// TIA Portal V20 export
// export: Created 2026-10-19T18:36:12.7338711Z, ExportSetting WithDefaults, DisplayName Totally Integrated Automation Portal, DisplayVersion V20 Update 6, DisplayName TIA Portal Openness, DisplayVersion V20 Update 6, DisplayName TIA Portal Version Control Interface, DisplayVersion V20 Update 6, DisplayName SINAMICS Startdrive Advanced, DisplayVersion V20 SP1, DisplayName SINAMICS Startdrive G130, G150, S120, S150, SINAMICS MV, G220, S200, S210, DisplayVersion V20 SP1, DisplayName SINAMICS Startdrive G110M, G120, G120C, G120D, G120P, G115D, DisplayVersion V20 SP1, DisplayName STEP 7 Professional, DisplayVersion V20 Update 6, DisplayName STEP 7 Safety, DisplayVersion V20 Update 2, DisplayName WinCC Basic/Comfort/Advanced, DisplayVersion V20 Update 6, DisplayName WinCC Unified, DisplayVersion V20 Update 6
FUNCTION "CNV_Order_FC" : Void   // FC46, SCL
{ S7_Optimized_Access := 'TRUE' }
VERSION : 0.1
// stored: AutoNumber true, IsIECCheckEnabled false, SetENOAutomatically false, UDAEnableTagReadback false
   VAR_INPUT
      i_Sys : UInt;
      Level : UInt;
      Tower : UInt;
      Transfer_From_To : Byte;
      Device : String;
      Task_Type : Int;
   END_VAR
   VAR_IN_OUT
      StepTable_0 : "OrderTable_UDT";
   END_VAR
   VAR_TEMP
      StrSys : String;
      StrLev : String;
      Concat1 : String;
      Concat2 : String;
      Source_Location : DInt;
      Destination_Location : DInt;
      Concat3 : String;
      Concat4 : String;
      StrSource : String;
      StrDestination : String;
   END_VAR
BEGIN
   #StrSys := UINT_TO_STRING(#i_Sys);

   // Remove "+"
   IF #StrSys[1] = '+' THEN
       #StrSys := RIGHT(IN := #StrSys, L := LEN(#StrSys) - 1);
   END_IF;

   #StrLev := UINT_TO_STRING(#Level);

   // Remove "+"
   IF #StrLev[1] = '+' THEN
       #StrLev := RIGHT(IN := #StrLev, L := LEN(#StrLev) - 1);
   END_IF;

   IF #Tower = 1 AND #Transfer_From_To = 1 THEN//EXTRACTOR TO CONVEYOR 1
       #StrSource := '120';
       #StrDestination := '100';
   ELSIF #Tower = 1 AND #Transfer_From_To = 2 THEN //CONVEYOR 1 TO EXTRACTOR
       #StrSource := '100';
       #StrDestination := '120';
   ELSIF #Tower = 2 AND #Transfer_From_To = 1 THEN //CONVEYOR 1 TO CONVEYOR 2
       #StrSource := '100';
       #StrDestination := '110';
   ELSIF #Tower = 2 AND #Transfer_From_To = 2 THEN //CONVEYOR 2 TO CONVEYOR 1
       #StrSource := '110';
       #StrDestination := '100';
   ELSIF #Tower = 0 AND #Transfer_From_To = 3 THEN //LOGISTEX TO EXTRACTOR
       #StrSource := '0';
       #StrDestination := '120';
   ELSIF #Tower = 0 AND #Transfer_From_To = 4 THEN // EXTRACTOR TO LOGISTEX
       #StrSource := '120';
       #StrDestination := '0';
   END_IF;

   // Build Source Location
   #Concat1 := CONCAT(IN1 := #StrSource, IN2 := #StrLev);
   #Concat2 := CONCAT(IN1 := #Concat1, IN2 := '0');
   #Source_Location := STRING_TO_DINT(IN := CONCAT(IN1 := #Concat2, IN2 := #StrSys));

   // Build Destinarion Location
   #Concat3 := CONCAT(IN1 := #StrDestination, IN2 := #StrLev);
   #Concat4 := CONCAT(IN1 := #Concat3, IN2 := '0');
   #Destination_Location := STRING_TO_DINT(IN := CONCAT(IN1 := #Concat4, IN2 := #StrSys));

   "Feed_Steptable_FC"(CurrentTime := "Time".CurrentLocalTime,
                       Task_Type := #Task_Type,
                       Source_Location := #Source_Location,
                       Destination_Location := #Destination_Location,
                       Shuttle_ID:=0,
                       StepTable := #StepTable_0);
END_FUNCTION
